Fanuc KAREL source: KA00067.KL

PROGRAM KA00067
%NOLOCKGROUP
VAR
  SRC: XYZWPR
  DST: XYZWPREXT
BEGIN
  SRC.X = 1.0
  DST = SRC
END KA00067
